(* IEC 61131-3 sources: llm-plc-st-eval/data/raw/gpt-4o/I2/few_shot, 3 files *)

(* ---- ejec_1.st ---- *)
```pascal
FUNCTION_BLOCK FB_Llenado
VAR_INPUT
    nivelAlto : BOOL; (* Sensor de nivel alto *)
    nivelBajo : BOOL; (* Sensor de nivel bajo *)
    btnInicio : BOOL; (* Botón de inicio del proceso *)
    btnParo : BOOL;   (* Botón de paro del proceso *)
END_VAR
VAR_OUTPUT
    vLlenado : BOOL;  (* Válvula de llenado *)
    motorMezcla : BOOL; (* Motor de mezcla *)
    vDescarga : BOOL; (* Válvula de descarga *)
END_VAR
VAR
    estado : INT := 0; (* Estado del proceso *)
    tMezcla : TON;     (* Temporizador para el motor de mezcla *)
END_VAR

(* Lógica del proceso de llenado por etapas *)
IF btnParo THEN
    (* Si se presiona el botón de paro, detener el proceso y resetear *)
    estado := 0;
    vLlenado := FALSE;
    motorMezcla := FALSE;
    vDescarga := FALSE;
ELSE
    CASE estado OF
        0: (* Estado de reposo *)
            IF btnInicio THEN
                estado := 1; (* Iniciar proceso de llenado *)
            END_IF;
        1: (* Llenado del tanque *)
            vLlenado := TRUE;
            IF nivelAlto THEN
                vLlenado := FALSE;
                estado := 2; (* Pasar al estado de mezcla *)
                tMezcla(IN := TRUE, PT := T#60S); (* Iniciar temporizador de mezcla *)
            END_IF;
        2: (* Mezcla del contenido *)
            motorMezcla := TRUE;
            tMezcla(IN := TRUE);
            IF tMezcla.Q THEN
                motorMezcla := FALSE;
                estado := 3; (* Pasar al estado de descarga *)
            END_IF;
        3: (* Descarga del tanque *)
            vDescarga := TRUE;
            IF nivelBajo THEN
                vDescarga := FALSE;
                estado := 0; (* Volver al estado de reposo *)
            END_IF;
    END_CASE;
END_IF;
END_FUNCTION_BLOCK
```

(* ---- ejec_2.st ---- *)
```pascal
FUNCTION_BLOCK FB_Llenado
VAR_INPUT
    nivelAlto : BOOL; (* Sensor de nivel alto *)
    nivelBajo : BOOL; (* Sensor de nivel bajo *)
    btnInicio : BOOL; (* Botón de inicio del proceso *)
    btnParo : BOOL;   (* Botón de paro de emergencia *)
END_VAR
VAR_OUTPUT
    vLlenado : BOOL;  (* Válvula de llenado *)
    motorMezcla : BOOL; (* Motor de mezcla *)
    vDescarga : BOOL; (* Válvula de descarga *)
END_VAR
VAR
    estado : INT := 0; (* Estado del proceso *)
    tMezcla : TON;     (* Temporizador para el motor de mezcla *)
END_VAR

(* Lógica de control del proceso de llenado por etapas *)
IF btnParo THEN
    (* Paro de emergencia: todas las salidas desactivadas y proceso en reposo *)
    estado := 0;
    vLlenado := FALSE;
    motorMezcla := FALSE;
    vDescarga := FALSE;
ELSIF btnInicio THEN
    CASE estado OF
        0: (* Estado de reposo *)
            IF btnInicio THEN
                estado := 1; (* Iniciar llenado *)
            END_IF;
        1: (* Llenado *)
            vLlenado := TRUE;
            IF nivelAlto THEN
                vLlenado := FALSE;
                estado := 2; (* Iniciar mezcla *)
                tMezcla(IN := TRUE, PT := T#60S);
            END_IF;
        2: (* Mezcla *)
            motorMezcla := tMezcla.Q;
            IF NOT tMezcla.Q THEN
                estado := 3; (* Iniciar descarga *)
            END_IF;
        3: (* Descarga *)
            vDescarga := TRUE;
            IF nivelBajo THEN
                vDescarga := FALSE;
                estado := 0; (* Volver a reposo *)
            END_IF;
    END_CASE;
END_IF;
END_FUNCTION_BLOCK
```

(* ---- ejec_3.st ---- *)
```pascal
FUNCTION_BLOCK FB_Llenado
VAR_INPUT
    nivelAlto : BOOL; (* Sensor de nivel alto *)
    nivelBajo : BOOL; (* Sensor de nivel bajo *)
    btnInicio : BOOL; (* Botón de inicio *)
    btnParo : BOOL; (* Botón de paro *)
END_VAR
VAR_OUTPUT
    vLlenado : BOOL; (* Válvula de llenado *)
    motorMezcla : BOOL; (* Motor de mezcla *)
    vDescarga : BOOL; (* Válvula de descarga *)
END_VAR
VAR
    estado : INT := 0; (* Estado del proceso *)
    tMezcla : TON; (* Temporizador para mezcla *)
END_VAR

(* Control del proceso de llenado por etapas *)
CASE estado OF
    0: (* Estado de reposo *)
        vLlenado := FALSE;
        motorMezcla := FALSE;
        vDescarga := FALSE;
        IF btnInicio THEN
            estado := 1; (* Iniciar llenado *)
        END_IF;
    1: (* Estado de llenado *)
        vLlenado := TRUE;
        IF nivelAlto THEN
            vLlenado := FALSE;
            tMezcla(IN := TRUE, PT := T#60S);
            estado := 2; (* Iniciar mezcla *)
        END_IF;
    2: (* Estado de mezcla *)
        motorMezcla := tMezcla.Q;
        IF NOT tMezcla.Q THEN
            motorMezcla := FALSE;
            estado := 3; (* Iniciar descarga *)
        END_IF;
    3: (* Estado de descarga *)
        vDescarga := TRUE;
        IF nivelBajo THEN
            vDescarga := FALSE;
            estado := 0; (* Volver a reposo *)
        END_IF;
END_CASE;

(* Manejo del botón de paro *)
IF btnParo THEN
    vLlenado := FALSE;
    motorMezcla := FALSE;
    vDescarga := FALSE;
    estado := 0; (* Volver a reposo *)
END_IF;
END_FUNCTION_BLOCK
```
